// TIA Portal V21 export
// export: Created 2026-11-10T07:02:24.8034991Z, ExportSetting WithDefaults, DisplayName Totally Integrated Automation Portal, DisplayVersion V21 Update 3, DisplayName STEP 7 Professional, DisplayVersion V21 Update 3, DisplayName STEP 7 Safety, DisplayVersion V21, DisplayName Tech WebApplication, DisplayVersion V21, DisplayName WinCC Basic/Comfort/Advanced, DisplayVersion V21 Update 3, DisplayName WinCC Unified, DisplayVersion V21 Update 3
FUNCTION "FC_SclMisc" : Void   // FC9, SCL
{ S7_Optimized_Access := 'TRUE' }
VERSION : 0.1
// stored: AutoNumber true, IsIECCheckEnabled false, SetENOAutomatically false, UDAEnableTagReadback false
   VAR_IN_OUT
      arr : Array[1..2, 1..2] of Int;
      arr3 : Array[0..1, 0..1, 0..1] of Int;
   END_VAR
   VAR_TEMP
      i : Int;
      d : DInt;
      "b" : Bool;
      v : Variant;
      "by" : Byte;
      w : Word;
      p : Int;
   END_VAR
BEGIN
   #by := PEEK(area := 16#84, dbNumber := 1, byteOffset := 0);
   POKE(area := 16#84, dbNumber := 1, byteOffset := 0, value := #by);
   #w := PEEK_WORD(area := 16#84, dbNumber := 1, byteOffset := 0);
   POKE(area := 16#84, dbNumber := 1, byteOffset := 0, value := #w);
   #b := PEEK_BOOL(area := 16#84, dbNumber := 1, byteOffset := 0, bitOffset := 1);
   #v := REF("DB_Global".iInt);
   #arr[1, 1] := 1;
   #arr3[0, 1, 0] := 3;
   #b := IS_ARRAY(#v);
   #i := CountOfElements(#v);
   #d := #i;
END_FUNCTION
